Fanuc KAREL source: kb00122.KL

-- PROVISIONAL review KL for V770-1; original PC SHA256 c9bca93751dc2da69a9184fd97bb057c772a2f85aa5e2eb54efaf7a02f287c3e
-- Incomplete behavior may be omitted. Consult companion uncertainty JSON. Do not deploy.
PROGRAM KB00122
%NOLOCKGROUP
BEGIN
  -- UNRESOLVED_PC offsets 5-14; opcodes 3F,75
  -- UNRESOLVED_PC offsets 19-26; opcodes 9D,23
  -- UNRESOLVED_PC offsets 31-49; opcodes 27,22,2A,22,31
  -- UNRESOLVED_PC offsets 54-58; opcodes 7F
END KB00122
